(* IEC 61131-3 sources: Caravan/Archiv/12-04-19/Stations/MachineControl/MachineControl/Network/Level_NET, 1 file *)

(* ---- ONE_Level_Net_Table.st ---- *)
#define OBJECTS_CONFIG

FUNCTION GLOBAL TAB ONE_Level_Net
-1$UINT, 0$UINT,
0$UINT, 0$UINT,

2$UDINT,
TO_UDINT(222137160), "Level_Class", 0$UINT, 0$UINT, 1$UINT,
TO_UDINT(912864977), "LevelFilter_Class", 0$UINT, 0$UINT, 1$UINT,

_NO_ATTR, TO_UDINT(4225112990), "LEVEL_CLASS1",

_NO_ATTR, TO_UDINT(1916691651), "LEVELFILTER_CLASS1",

//Internal connections
0$UDINT,
0$UDINT,
0$UDINT,
2$UDINT,
TO_UDINT(0), "PositionInput_X_C", TO_UDINT(1), "X_Out_S",
TO_UDINT(0), "PositionInput_Y_C", TO_UDINT(1), "Y_Out_S",

//Initialization values
0$UDINT,
1$UDINT,
TO_UDINT(1), "Y_IN_C", TO_UDINT(0),//|Level_Net.LevelFilter_Class1.Y_IN_C;

//Symbolic initialization values
0$UDINT,
0$UDINT,

//Initialization of string values
0$UDINT,
0$UDINT,

//Configuration of tasks (RealTime, Cyclic, Background)
0$UDINT,
0$UDINT,

0$UDINT,
2$UDINT,
TO_UDINT(0), (50)$UDINT, 4194303$DINT, 	//LEVEL_CLASS1
TO_UDINT(1), (10)$UDINT, 4194303$DINT, 	//LEVELFILTER_CLASS1

0$UDINT,
0$UDINT,

//External connections
0$UDINT,
2$UDINT,
TO_UDINT(1), "X_IN_C", C_DIR, TO_UDINT(46500714), "AI0751","AI2",
TO_UDINT(1), "Y_IN_C", C_DIR, TO_UDINT(46500714), "AI0751","AI3",

//Magic internal connections
0$UDINT,
0$UDINT,

//Configuration of timeslots of tasks (RealTime, Cyclic)
#ifdef __LSLLDR_TIMESLOTS__
0$UDINT,
0$UDINT,

0$UDINT,
0$UDINT,

#endif //__LSLLDR_TIMESLOTS__

//MultiMaster connections
#ifdef __LSLLDR_MULTIMASTER__
0$UDINT,
0$UDINT,
#endif //__LSLLDR_MULTIMASTER__

//Configuration for task ID (RealTime, CyclicTime)
#ifdef __LSLLDR_TASKID__
"\\\\TASKS2  "
0$UDINT,
0$UDINT,

0$UDINT,
2$UDINT,
(0)$UDINT, 	//LEVEL_CLASS1
(0)$UDINT, 	//LEVELFILTER_CLASS1

0$UDINT,
0$UDINT,

#endif //__LSLLDR_TASKID__

END_FUNCTION
